// TIA Portal V19 export
TYPE "EM_Input"
   STRUCT
      Start : Bool;   // Comando por flanco: inicia desde Idle o reanuda desde Held
      Stop : Bool;   // Comando por flanco: detiene de forma ordenada
      Hold : Bool;   // Comando por flanco: pausa la ejecuciÃ³n
      Abort : Bool;   // Comando por flanco: aborta (mÃ¡xima prioridad)
      Reset : Bool;   // Comando por flanco: limpia fallos y regresa a Idle
      Manual : Bool;
      Auto : Bool;
      Maintenance : Bool;
   END_STRUCT;
END_TYPE
